// TIA Portal V20 export
TYPE "WT2_Vr_Befehl_UDT"
   STRUCT
      iHandshake : Int;
      Befehl : Struct
         iID : Int;
         iParam : Int;
      END_STRUCT;
      Param : Struct
         diID : DInt;
         diValue : DInt;
         iDiv : Int;
         byEditKonfigSet : Byte;
         byReserve : Byte;
         diReserve2 : DInt;
      END_STRUCT;
      FernVorgabeDig : Struct
         bFreigabeNiveauregAbsch : Bool;
         bSollwertumschAB : Bool;
         b222_Reserve : Bool;
         b223_Reserve : Bool;
         b224_Reserve : Bool;
         b225_Reserve : Bool;
         b226_Reserve : Bool;
         b227_Reserve : Bool;
         by23_Reserve : Byte;
      END_STRUCT;
      rFernSollwert : Real;
      rReserveReal : Array[0..3] of Real;
   END_STRUCT;
END_TYPE
